(* IEC 61131-3 sources: codesys-framework/txt/application/WeVe Core (library)/60 Event/FB_Event/Private, 2 files *)

(* ---- FillPlaceholders.method.st ---- *)
// Vervangt %0..%9 in sTemplate door scPayload.asPayload[0..9].
// Een '%' die niet gevolgd wordt door een cijfer blijft staan (bv. '50 %').
METHOD PRIVATE FillPlaceholders : STRING(GVL_Logger.cMaxMessageLength)
VAR_INPUT
	sTemplate 		: STRING(GVL_Logger.cMaxMessageLength);
	scPayload 		: SC_EventPayload;
END_VAR
VAR
	sResult 		: STRING(GVL_Logger.cMaxMessageLength);
	sRest 			: STRING(GVL_Logger.cMaxMessageLength);
	iPos 			: INT;		// positie van '%' in sRest, 1-gebaseerd (FIND)
	byNext 			: BYTE;		// teken na '%'
END_VAR

// --- BEGIN IMPLEMENTATION ---

sResult := '';
sRest := sTemplate;
iPos := FIND(sRest, '%');

WHILE iPos > 0 DO

	// Alles voor de '%' overnemen
	sResult := CONCAT(sResult, LEFT(sRest, iPos - 1));

	// sRest[i] is 0-gebaseerd: sRest[iPos] is het teken na '%' (0 als '%' het laatste teken is)
	byNext := sRest[iPos];

	IF byNext >= 16#30 AND byNext <= 16#39 THEN
		sResult := CONCAT(sResult, scPayload.asPayload[byNext - 16#30]);
		sRest := RIGHT(sRest, LEN(sRest) - iPos - 1);
	ELSE
		sResult := CONCAT(sResult, '%');
		sRest := RIGHT(sRest, LEN(sRest) - iPos);
	END_IF

	iPos := FIND(sRest, '%');

END_WHILE

FillPlaceholders := CONCAT(sResult, sRest);

(* ---- WriteLog.method.st ---- *)
// Bouwt de logregel op en geeft ze door aan de logger.
//   '<level> [<overgang>] | <id> | <subMachine>.<subMachineId> | <boodschap>'
// sTransition = '' voor een eenmalige melding.
// TRUE = gelogd. FALSE = geen logger of buffer vol.
METHOD PRIVATE WriteLog : BOOL
VAR_INPUT
	sTransition 	: STRING(20);
	scPayload 		: SC_EventPayload;
END_VAR
VAR
	sLine 			: STRING(GVL_Logger.cMaxMessageLength);
END_VAR

// --- BEGIN IMPLEMENTATION ---

IF _fbLogger = 0 THEN
	WriteLog := FALSE;
	RETURN;
END_IF

sLine := F_EventLevelToText(_scConfig.eEventLevel);

IF sTransition <> '' THEN
	sLine := CONCAT(sLine, ' ');
	sLine := CONCAT(sLine, sTransition);
END_IF

sLine := CONCAT(sLine, ' | ');
sLine := CONCAT(sLine, UDINT_TO_STRING(_scConfig.udiEventId));
sLine := CONCAT(sLine, ' | ');
sLine := CONCAT(sLine, USINT_TO_STRING(_scConfig.nSubMachine));
sLine := CONCAT(sLine, '.');
sLine := CONCAT(sLine, USINT_TO_STRING(_scConfig.nSubMachineId));
sLine := CONCAT(sLine, ' | ');
sLine := CONCAT(sLine, FillPlaceholders(sTemplate := _scConfig.sMessage, scPayload := scPayload));

WriteLog := _fbLogger.LogEvent(scEvent := _scConfig, scPayload := scPayload, sMessage := sLine);
